{attribute 'qualified_only'}
{attribute 'strict'}
{attribute 'to_string'}
TYPE E_PolarIIChamberCycleControl :
(
	None := 0,
	Start := 1,
	End := 2
) UINT;
END_TYPE

(* stored: Version 1.1.0.1, ProductVersion 3.1.4026.18
   DUT E_PolarIIChamberCycleControl: Id {14000000-0000-0000-0000-000000000005} *)
